// Mitsubishi GX Works2 project: 미니프로젝트 합본   PLC: Q03UDV

PROGRAM MAIN
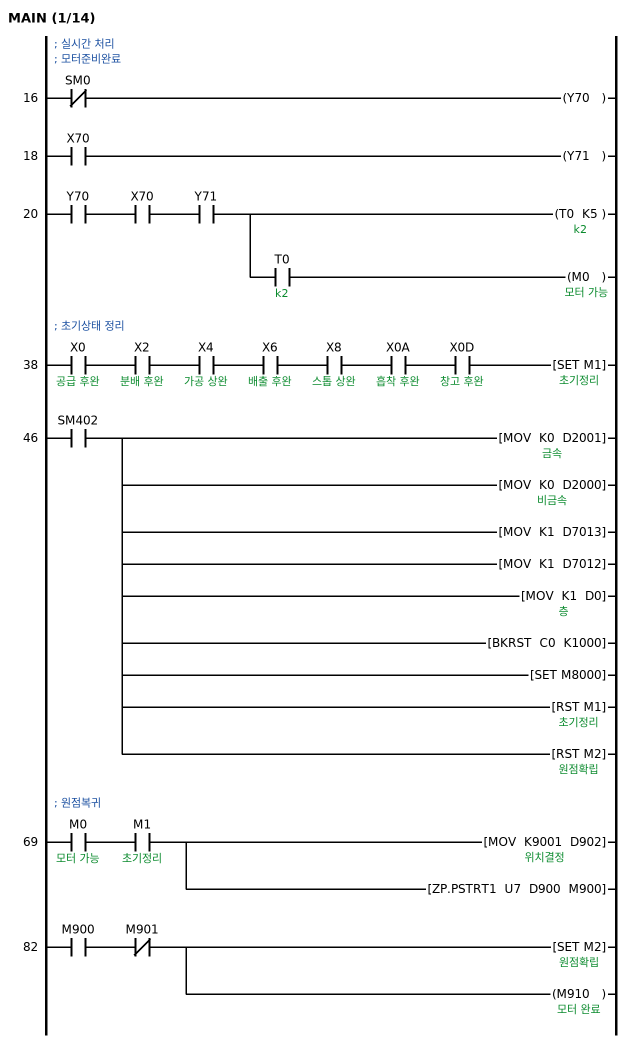
; 실시간 처리
; 모터준비완료
16    LDI     SM0
      OUT     Y70
18    LD      X70
      OUT     Y71
20    LD      Y70
      AND     X70
      AND     Y71
      OUT     T0 K5  ; k2
      AND     T0  ; k2
      OUT     M0  ; 모터 가능
; 초기상태 정리
38    LD      X0  ; 공급 후완
      AND     X2  ; 분배 후완
      AND     X4  ; 가공 상완
      AND     X6  ; 배출 후완
      AND     X8  ; 스톱 상완
      AND     X0A  ; 흡착 후완
      AND     X0D  ; 창고 후완
      SET     M1  ; 초기정리
46    LD      SM402
      MOV     K0 D2001  ; 금속
      MOV     K0 D2000  ; 비금속
      MOV     K1 D7013
      MOV     K1 D7012
      MOV     K1 D0  ; 층
      BKRST   C0 K1000
      SET     M8000
      RST     M1  ; 초기정리
      RST     M2  ; 원점확립
; 원점복귀
69    LD      M0  ; 모터 가능
      AND     M1  ; 초기정리
      MOV     K9001 D902  ; 위치결정
      ZP.PSTRT1 U7 D900 M900
82    LD      M900
      ANI     M901
      SET     M2  ; 원점확립
      OUT     M910  ; 모터 완료
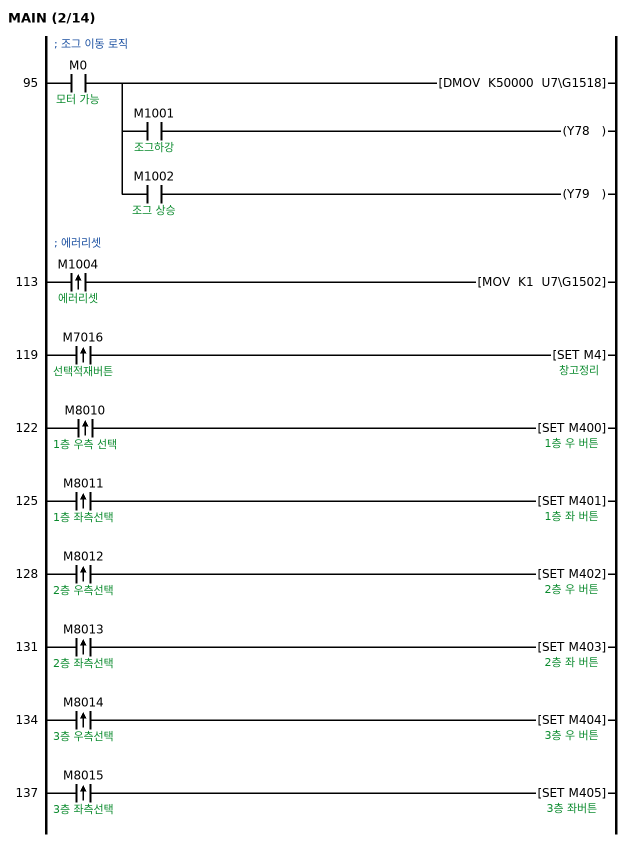
; 조그 이동 로직
95    LD      M0  ; 모터 가능
      DMOV    K50000 U7\G1518
      MPS
      AND     M1001  ; 조그하강
      OUT     Y78
      MPP
      AND     M1002  ; 조그 상승
      OUT     Y79
; 에러리셋
113   LDP     M1004  ; 에러리셋
      MOV     K1 U7\G1502
119   LDP     M7016  ; 선택적재버튼
      SET     M4  ; 창고정리
122   LDP     M8010  ; 1층 우측 선택
      SET     M400  ; 1층 우 버튼
125   LDP     M8011  ; 1층 좌측선택
      SET     M401  ; 1층 좌 버튼
128   LDP     M8012  ; 2층 우측선택
      SET     M402  ; 2층 우 버튼
131   LDP     M8013  ; 2층 좌측선택
      SET     M403  ; 2층 좌 버튼
134   LDP     M8014  ; 3층 우측선택
      SET     M404  ; 3층 우 버튼
137   LDP     M8015  ; 3층 좌측선택
      SET     M405  ; 3층 좌버튼
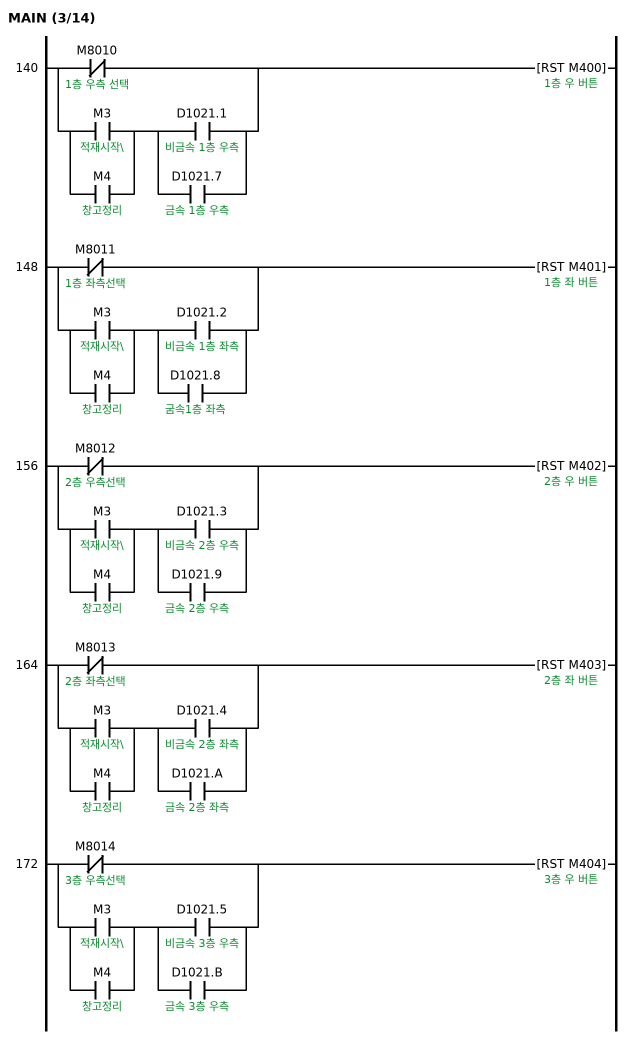
140   LDI     M8010  ; 1층 우측 선택
      LD      M3  ; 적재시작\
      OR      M4  ; 창고정리
      LD      D1021.1  ; 비금속 1층 우측
      OR      D1021.7  ; 금속 1층 우측
      ANB
      ORB
      RST     M400  ; 1층 우 버튼
148   LDI     M8011  ; 1층 좌측선택
      LD      M3  ; 적재시작\
      OR      M4  ; 창고정리
      LD      D1021.2  ; 비금속 1층 좌측
      OR      D1021.8  ; 굼속1층 좌측
      ANB
      ORB
      RST     M401  ; 1층 좌 버튼
156   LDI     M8012  ; 2층 우측선택
      LD      M3  ; 적재시작\
      OR      M4  ; 창고정리
      LD      D1021.3  ; 비금속 2층 우측
      OR      D1021.9  ; 금속 2층 우측
      ANB
      ORB
      RST     M402  ; 2층 우 버튼
164   LDI     M8013  ; 2층 좌측선택
      LD      M3  ; 적재시작\
      OR      M4  ; 창고정리
      LD      D1021.4  ; 비금속 2층 좌측
      OR      D1021.A  ; 금속 2층 좌측
      ANB
      ORB
      RST     M403  ; 2층 좌 버튼
172   LDI     M8014  ; 3층 우측선택
      LD      M3  ; 적재시작\
      OR      M4  ; 창고정리
      LD      D1021.5  ; 비금속 3층 우측
      OR      D1021.B  ; 금속 3층 우측
      ANB
      ORB
      RST     M404  ; 3층 우 버튼
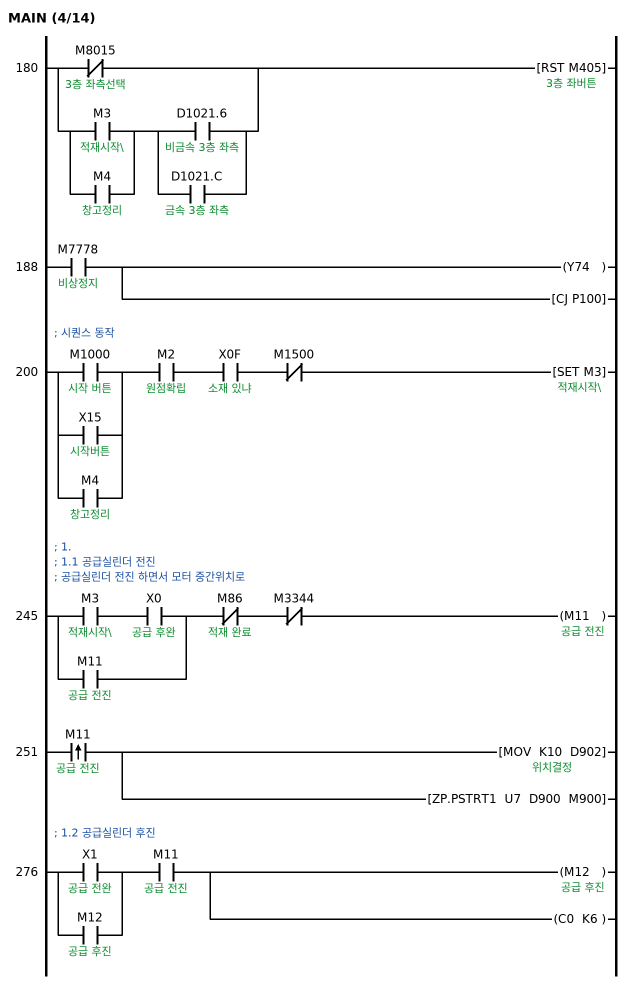
180   LDI     M8015  ; 3층 좌측선택
      LD      M3  ; 적재시작\
      OR      M4  ; 창고정리
      LD      D1021.6  ; 비금속 3층 좌측
      OR      D1021.C  ; 금속 3층 좌측
      ANB
      ORB
      RST     M405  ; 3층 좌버튼
188   LD      M7778  ; 비상정지
      OUT     Y74
      CJ      P100
; 시퀀스 동작
200   LD      M1000  ; 시작 버튼
      OR      X15  ; 시작버튼
      OR      M4  ; 창고정리
      AND     M2  ; 원점확립
      AND     X0F  ; 소재 있냐
      ANI     M1500
      SET     M3  ; 적재시작\
; 1.
; 1.1 공급실린더 전진
; 공급실린더 전진 하면서 모터 중간위치로
245   LD      M3  ; 적재시작\
      AND     X0  ; 공급 후완
      OR      M11  ; 공급 전진
      ANI     M86  ; 적재 완료
      ANI     M3344
      OUT     M11  ; 공급 전진
251   LDP     M11  ; 공급 전진
      MOV     K10 D902
      ZP.PSTRT1 U7 D900 M900
; 1.2 공급실린더 후진
276   LD      X1  ; 공급 전완
      OR      M12  ; 공급 후진
      AND     M11  ; 공급 전진
      OUT     M12  ; 공급 후진
      OUT     C0 K6
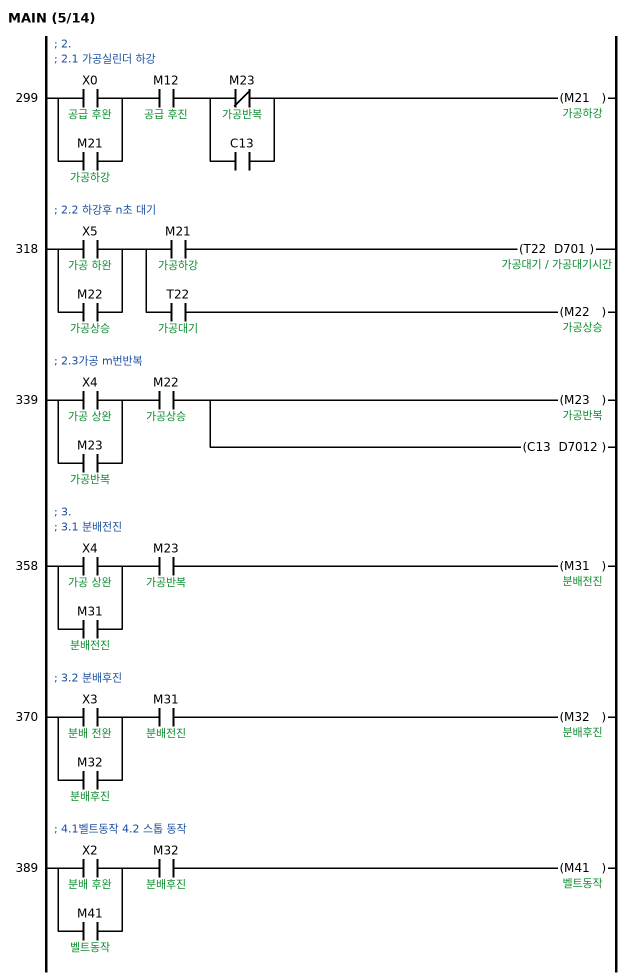
; 2.
; 2.1 가공실린더 하강
299   LD      X0  ; 공급 후완
      OR      M21  ; 가공하강
      AND     M12  ; 공급 후진
      LDI     M23  ; 가공반복
      OR      C13
      ANB
      OUT     M21  ; 가공하강
; 2.2 하강후 n초 대기
318   LD      X5  ; 가공 하완
      OR      M22  ; 가공상승
      MPS
      AND     M21  ; 가공하강
      OUT     T22 D701  ; 가공대기 / 가공대기시간
      MPP
      AND     T22  ; 가공대기
      OUT     M22  ; 가공상승
; 2.3가공 m번반복
339   LD      X4  ; 가공 상완
      OR      M23  ; 가공반복
      AND     M22  ; 가공상승
      OUT     M23  ; 가공반복
      OUT     C13 D7012
; 3.
; 3.1 분배전진
358   LD      X4  ; 가공 상완
      OR      M31  ; 분배전진
      AND     M23  ; 가공반복
      OUT     M31  ; 분배전진
; 3.2 분배후진
370   LD      X3  ; 분배 전완
      OR      M32  ; 분배후진
      AND     M31  ; 분배전진
      OUT     M32  ; 분배후진
; 4.1벨트동작 4.2 스톱 동작
389   LD      X2  ; 분배 후완
      OR      M41  ; 벨트동작
      AND     M32  ; 분배후진
      OUT     M41  ; 벨트동작
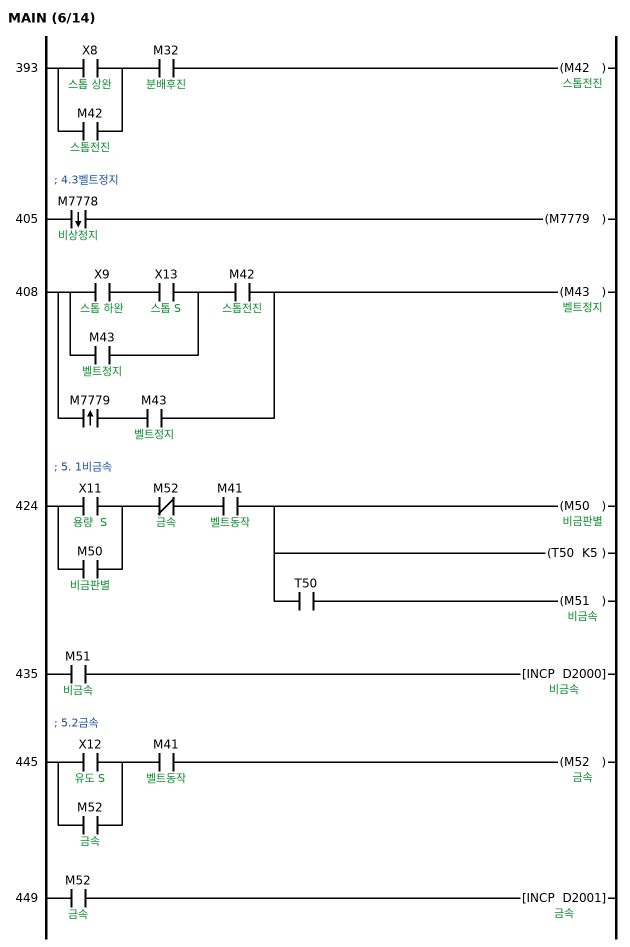
393   LD      X8  ; 스톱 상완
      OR      M42  ; 스톱전진
      AND     M32  ; 분배후진
      OUT     M42  ; 스톱전진
; 4.3벨트정지
405   LDF     M7778  ; 비상정지
      OUT     M7779
408   LD      X9  ; 스톱 하완
      AND     X13  ; 스톱 S
      OR      M43  ; 벨트정지
      AND     M42  ; 스톱전진
      LDP     M7779
      AND     M43  ; 벨트정지
      ORB
      OUT     M43  ; 벨트정지
; 5. 1비금속
424   LD      X11  ; 용량  S
      OR      M50  ; 비금판별
      ANI     M52  ; 금속
      AND     M41  ; 벨트동작
      OUT     M50  ; 비금판별
      OUT     T50 K5
      AND     T50
      OUT     M51  ; 비금속
435   LD      M51  ; 비금속
      INCP    D2000
; 5.2금속
445   LD      X12  ; 유도 S
      OR      M52  ; 금속
      AND     M41  ; 벨트동작
      OUT     M52  ; 금속
449   LD      M52  ; 금속
      INCP    D2001
      P100
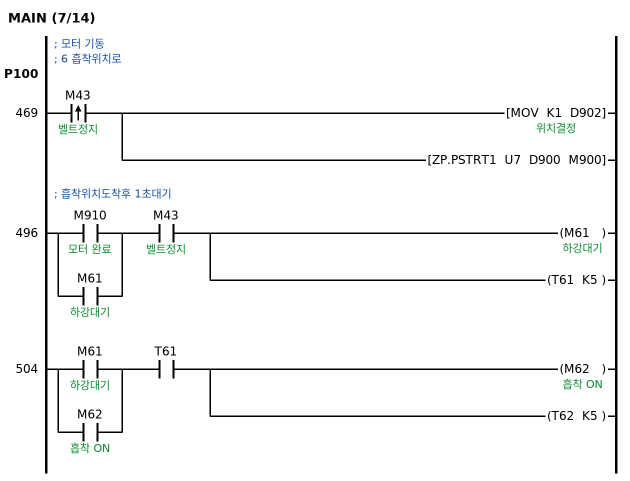
; 모터 기동
; 6 흡착위치로
469   LDP     M43  ; 벨트정지
      MOV     K1 D902
      ZP.PSTRT1 U7 D900 M900
; 흡착위치도착후 1초대기
496   LD      M910  ; 모터 완료
      OR      M61  ; 하강대기
      AND     M43  ; 벨트정지
      OUT     M61  ; 하강대기
      OUT     T61 K5
504   LD      M61  ; 하강대기
      OR      M62  ; 흡착 ON
      AND     T61
      OUT     M62  ; 흡착 ON
      OUT     T62 K5
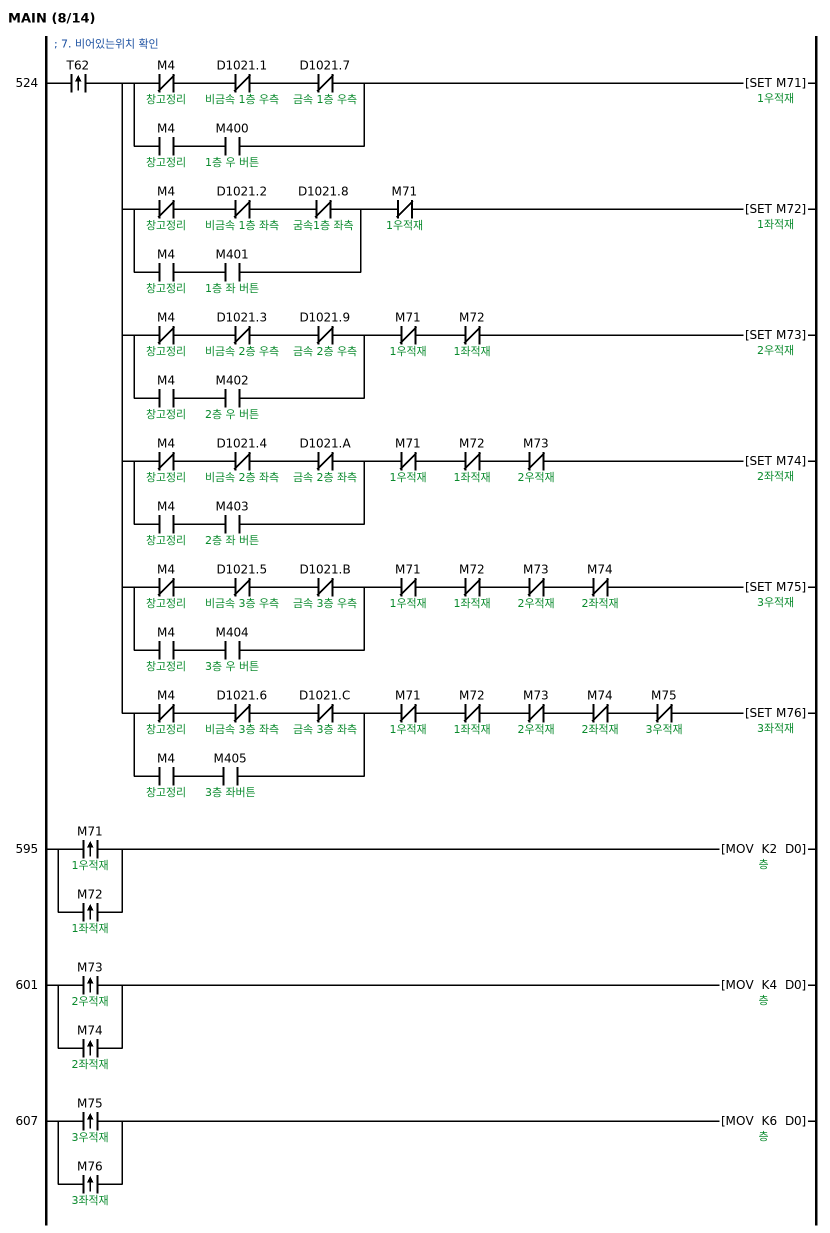
; 7. 비어있는위치 확인
524   LDP     T62
      MPS
      LDI     M4  ; 창고정리
      ANI     D1021.1  ; 비금속 1층 우측
      ANI     D1021.7  ; 금속 1층 우측
      LD      M4  ; 창고정리
      AND     M400  ; 1층 우 버튼
      ORB
      ANB
      SET     M71  ; 1우적재
      MRD
      LDI     M4  ; 창고정리
      ANI     D1021.2  ; 비금속 1층 좌측
      ANI     D1021.8  ; 굼속1층 좌측
      LD      M4  ; 창고정리
      AND     M401  ; 1층 좌 버튼
      ORB
      ANB
      ANI     M71  ; 1우적재
      SET     M72  ; 1좌적재
      MRD
      LDI     M4  ; 창고정리
      ANI     D1021.3  ; 비금속 2층 우측
      ANI     D1021.9  ; 금속 2층 우측
      LD      M4  ; 창고정리
      AND     M402  ; 2층 우 버튼
      ORB
      ANB
      ANI     M71  ; 1우적재
      ANI     M72  ; 1좌적재
      SET     M73  ; 2우적재
      MRD
      LDI     M4  ; 창고정리
      ANI     D1021.4  ; 비금속 2층 좌측
      ANI     D1021.A  ; 금속 2층 좌측
      LD      M4  ; 창고정리
      AND     M403  ; 2층 좌 버튼
      ORB
      ANB
      ANI     M71  ; 1우적재
      ANI     M72  ; 1좌적재
      ANI     M73  ; 2우적재
      SET     M74  ; 2좌적재
      MRD
      LDI     M4  ; 창고정리
      ANI     D1021.5  ; 비금속 3층 우측
      ANI     D1021.B  ; 금속 3층 우측
      LD      M4  ; 창고정리
      AND     M404  ; 3층 우 버튼
      ORB
      ANB
      ANI     M71  ; 1우적재
      ANI     M72  ; 1좌적재
      ANI     M73  ; 2우적재
      ANI     M74  ; 2좌적재
      SET     M75  ; 3우적재
      MPP
      LDI     M4  ; 창고정리
      ANI     D1021.6  ; 비금속 3층 좌측
      ANI     D1021.C  ; 금속 3층 좌측
      LD      M4  ; 창고정리
      AND     M405  ; 3층 좌버튼
      ORB
      ANB
      ANI     M71  ; 1우적재
      ANI     M72  ; 1좌적재
      ANI     M73  ; 2우적재
      ANI     M74  ; 2좌적재
      ANI     M75  ; 3우적재
      SET     M76  ; 3좌적재
595   LDP     M71  ; 1우적재
      ORP     M72  ; 1좌적재
      MOV     K2 D0
601   LDP     M73  ; 2우적재
      ORP     M74  ; 2좌적재
      MOV     K4 D0
607   LDP     M75  ; 3우적재
      ORP     M76  ; 3좌적재
      MOV     K6 D0
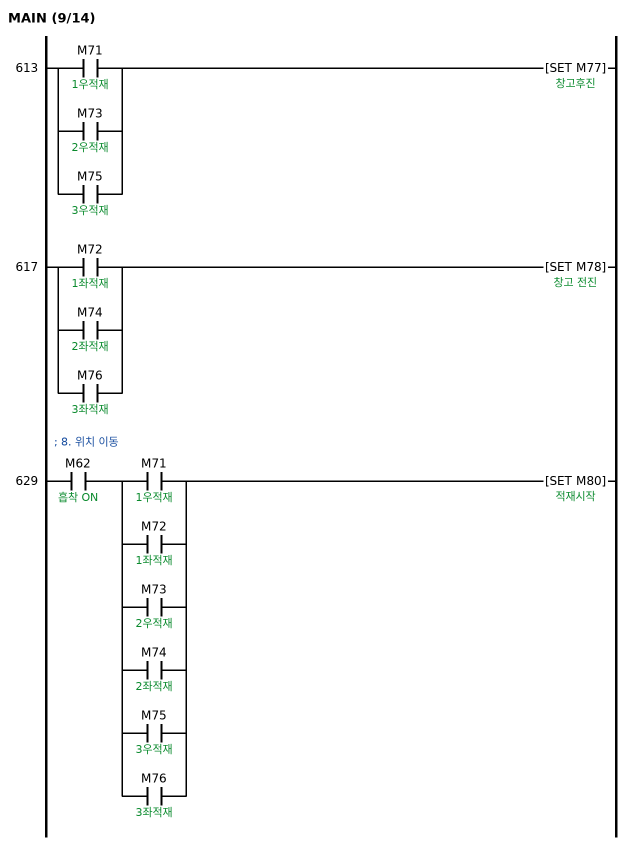
613   LD      M71  ; 1우적재
      OR      M73  ; 2우적재
      OR      M75  ; 3우적재
      SET     M77  ; 창고후진
617   LD      M72  ; 1좌적재
      OR      M74  ; 2좌적재
      OR      M76  ; 3좌적재
      SET     M78  ; 창고 전진
; 8. 위치 이동
629   LD      M62  ; 흡착 ON
      LD      M71  ; 1우적재
      OR      M72  ; 1좌적재
      OR      M73  ; 2우적재
      OR      M74  ; 2좌적재
      OR      M75  ; 3우적재
      OR      M76  ; 3좌적재
      ANB
      SET     M80  ; 적재시작
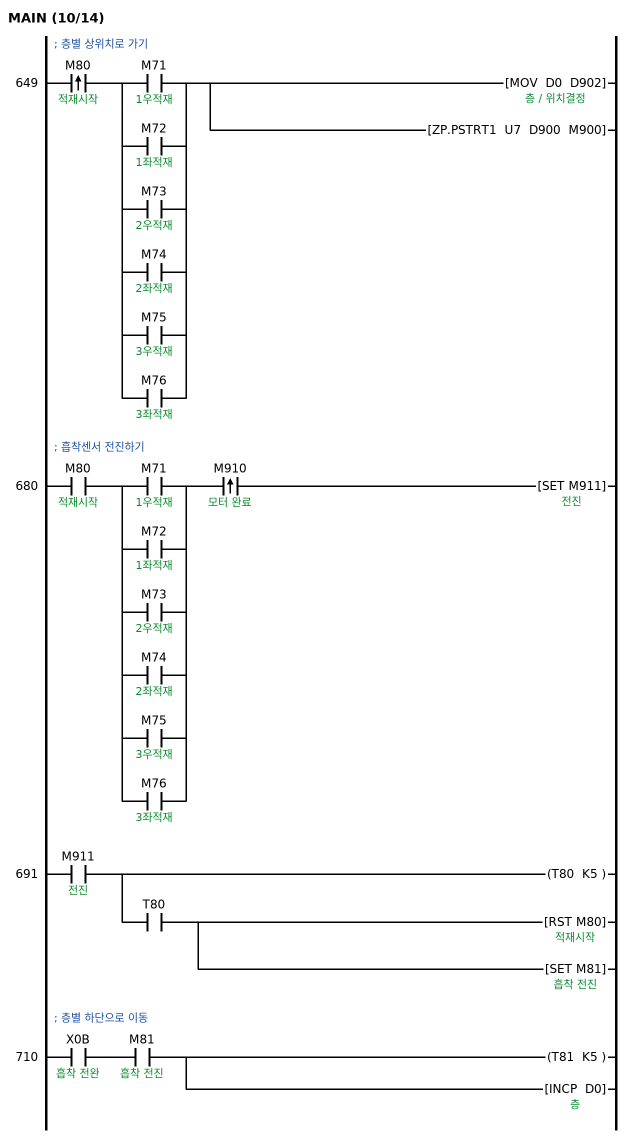
; 층별 상위치로 가기
649   LDP     M80  ; 적재시작
      LD      M71  ; 1우적재
      OR      M72  ; 1좌적재
      OR      M73  ; 2우적재
      OR      M74  ; 2좌적재
      OR      M75  ; 3우적재
      OR      M76  ; 3좌적재
      ANB
      MOV     D0 D902
      ZP.PSTRT1 U7 D900 M900
; 흡착센서 전진하기
680   LD      M80  ; 적재시작
      LD      M71  ; 1우적재
      OR      M72  ; 1좌적재
      OR      M73  ; 2우적재
      OR      M74  ; 2좌적재
      OR      M75  ; 3우적재
      OR      M76  ; 3좌적재
      ANB
      ANDP    M910  ; 모터 완료
      SET     M911  ; 전진
691   LD      M911  ; 전진
      OUT     T80 K5
      AND     T80
      RST     M80  ; 적재시작
      SET     M81  ; 흡착 전진
; 층별 하단으로 이동
710   LD      X0B  ; 흡착 전완
      AND     M81  ; 흡착 전진
      OUT     T81 K5
      INCP    D0
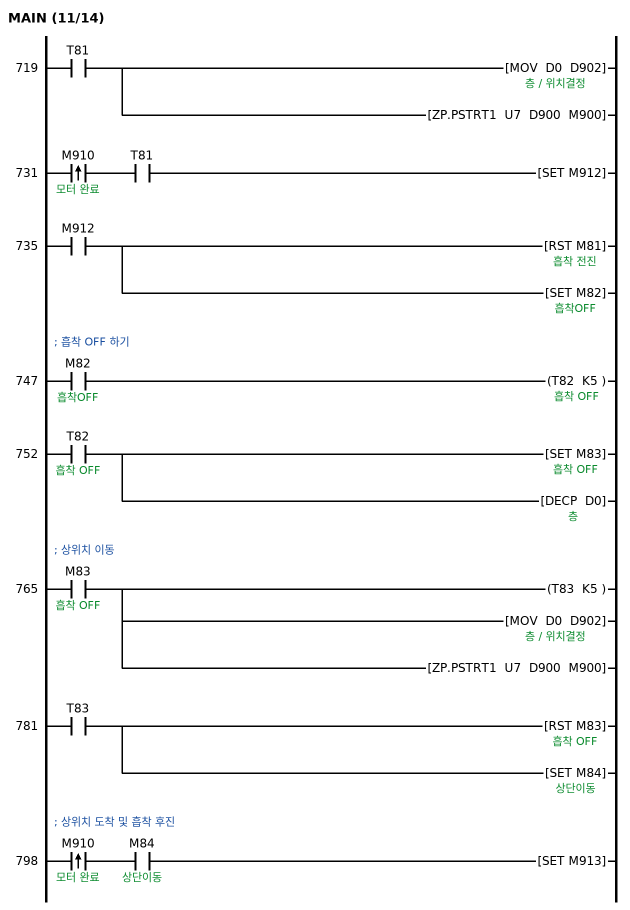
719   LD      T81
      MOV     D0 D902
      ZP.PSTRT1 U7 D900 M900
731   LDP     M910  ; 모터 완료
      AND     T81
      SET     M912
735   LD      M912
      RST     M81  ; 흡착 전진
      SET     M82  ; 흡착OFF
; 흡착 OFF 하기
747   LD      M82  ; 흡착OFF
      OUT     T82 K5  ; 흡착 OFF
752   LD      T82  ; 흡착 OFF
      SET     M83  ; 흡착 OFF
      DECP    D0
; 상위치 이동
765   LD      M83  ; 흡착 OFF
      OUT     T83 K5
      MOV     D0 D902
      ZP.PSTRT1 U7 D900 M900
781   LD      T83
      RST     M83  ; 흡착 OFF
      SET     M84  ; 상단이동
; 상위치 도착 및 흡착 후진
798   LDP     M910  ; 모터 완료
      AND     M84  ; 상단이동
      SET     M913
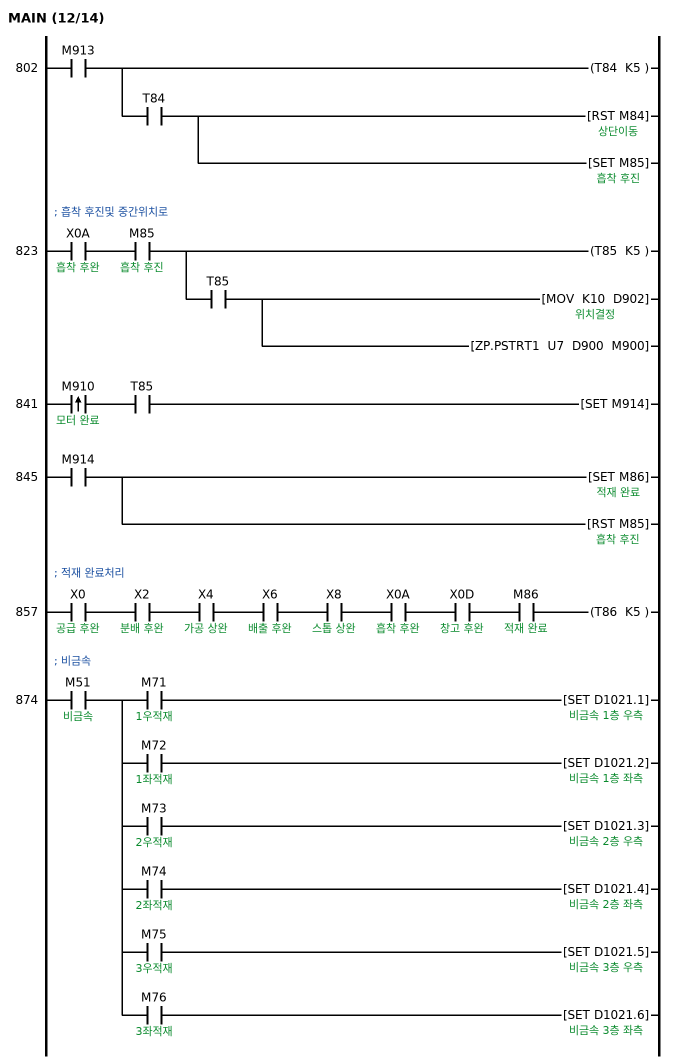
802   LD      M913
      OUT     T84 K5
      AND     T84
      RST     M84  ; 상단이동
      SET     M85  ; 흡착 후진
; 흡착 후진및 중간위치로
823   LD      X0A  ; 흡착 후완
      AND     M85  ; 흡착 후진
      OUT     T85 K5
      AND     T85
      MOV     K10 D902
      ZP.PSTRT1 U7 D900 M900
841   LDP     M910  ; 모터 완료
      AND     T85
      SET     M914
845   LD      M914
      SET     M86  ; 적재 완료
      RST     M85  ; 흡착 후진
; 적재 완료처리
857   LD      X0  ; 공급 후완
      AND     X2  ; 분배 후완
      AND     X4  ; 가공 상완
      AND     X6  ; 배출 후완
      AND     X8  ; 스톱 상완
      AND     X0A  ; 흡착 후완
      AND     X0D  ; 창고 후완
      AND     M86  ; 적재 완료
      OUT     T86 K5
; 비금속
874   LD      M51  ; 비금속
      MPS
      AND     M71  ; 1우적재
      SET     D1021.1  ; 비금속 1층 우측
      MRD
      AND     M72  ; 1좌적재
      SET     D1021.2  ; 비금속 1층 좌측
      MRD
      AND     M73  ; 2우적재
      SET     D1021.3  ; 비금속 2층 우측
      MRD
      AND     M74  ; 2좌적재
      SET     D1021.4  ; 비금속 2층 좌측
      MRD
      AND     M75  ; 3우적재
      SET     D1021.5  ; 비금속 3층 우측
      MPP
      AND     M76  ; 3좌적재
      SET     D1021.6  ; 비금속 3층 좌측
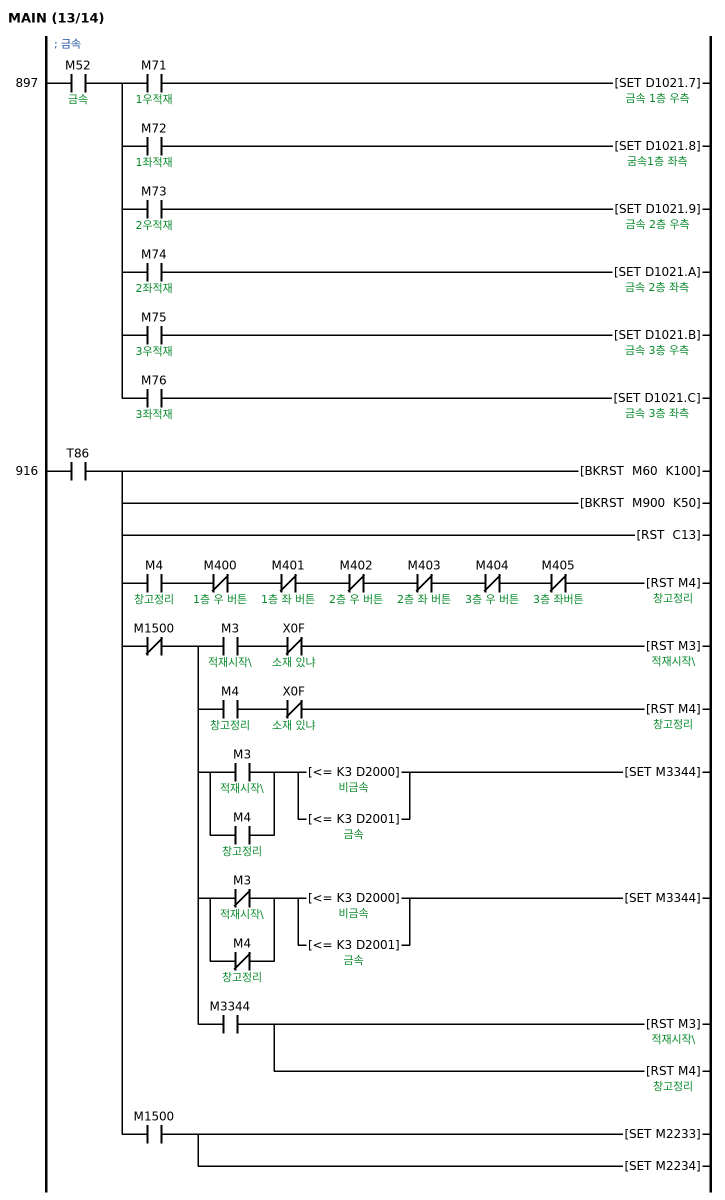
; 금속
897   LD      M52  ; 금속
      MPS
      AND     M71  ; 1우적재
      SET     D1021.7  ; 금속 1층 우측
      MRD
      AND     M72  ; 1좌적재
      SET     D1021.8  ; 굼속1층 좌측
      MRD
      AND     M73  ; 2우적재
      SET     D1021.9  ; 금속 2층 우측
      MRD
      AND     M74  ; 2좌적재
      SET     D1021.A  ; 금속 2층 좌측
      MRD
      AND     M75  ; 3우적재
      SET     D1021.B  ; 금속 3층 우측
      MPP
      AND     M76  ; 3좌적재
      SET     D1021.C  ; 금속 3층 좌측
916   LD      T86
      BKRST   M60 K100
      BKRST   M900 K50
      RST     C13
      MPS
      AND     M4  ; 창고정리
      ANI     M400  ; 1층 우 버튼
      ANI     M401  ; 1층 좌 버튼
      ANI     M402  ; 2층 우 버튼
      ANI     M403  ; 2층 좌 버튼
      ANI     M404  ; 3층 우 버튼
      ANI     M405  ; 3층 좌버튼
      RST     M4  ; 창고정리
      MRD
      ANI     M1500
      MPS
      AND     M3  ; 적재시작\
      ANI     X0F  ; 소재 있냐
      RST     M3  ; 적재시작\
      MRD
      AND     M4  ; 창고정리
      ANI     X0F  ; 소재 있냐
      RST     M4  ; 창고정리
      MRD
      LD      M3  ; 적재시작\
      OR      M4  ; 창고정리
      ANB
      LD<=    K3 D2000  ; 비금속
      OR<=    K3 D2001  ; 금속
      ANB
      SET     M3344
      MRD
      LDI     M3  ; 적재시작\
      ORI     M4  ; 창고정리
      ANB
      LD<=    K3 D2000  ; 비금속
      OR<=    K3 D2001  ; 금속
      ANB
      SET     M3344
      MPP
      AND     M3344
      RST     M3  ; 적재시작\
      RST     M4  ; 창고정리
      MPP
      AND     M1500
      SET     M2233
      SET     M2234
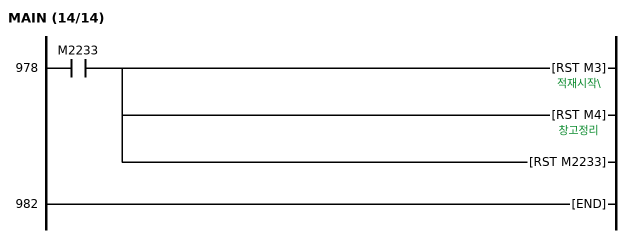
978   LD      M2233
      RST     M3  ; 적재시작\
      RST     M4  ; 창고정리
      RST     M2233
982   END
END_PROGRAM

PROGRAM OUTPUT
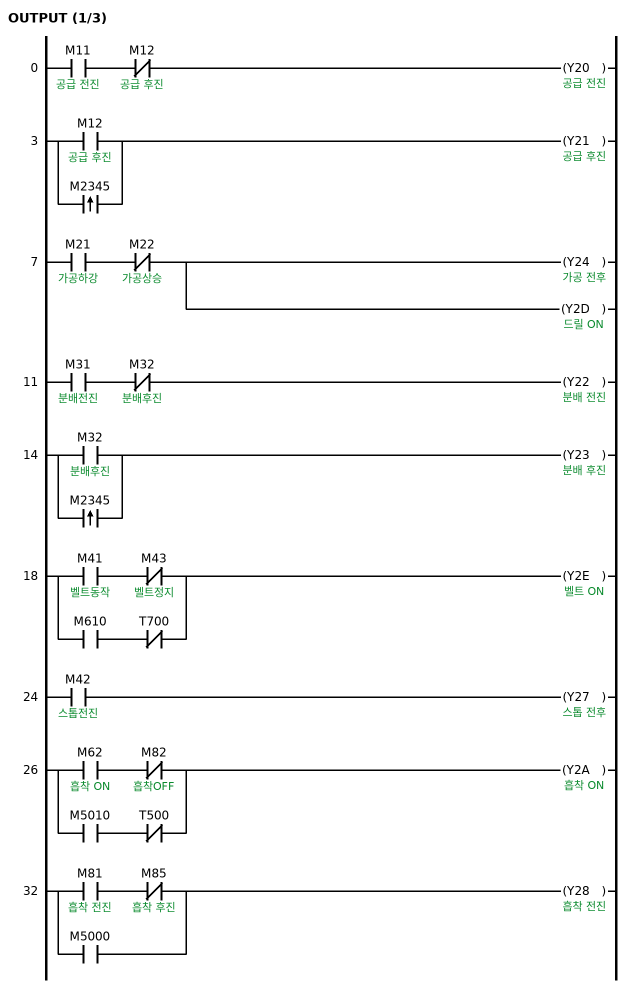
0     LD      M11  ; 공급 전진
      ANI     M12  ; 공급 후진
      OUT     Y20  ; 공급 전진
3     LD      M12  ; 공급 후진
      ORP     M2345
      OUT     Y21  ; 공급 후진
7     LD      M21  ; 가공하강
      ANI     M22  ; 가공상승
      OUT     Y24  ; 가공 전후
      OUT     Y2D  ; 드릴 ON
11    LD      M31  ; 분배전진
      ANI     M32  ; 분배후진
      OUT     Y22  ; 분배 전진
14    LD      M32  ; 분배후진
      ORP     M2345
      OUT     Y23  ; 분배 후진
18    LD      M41  ; 벨트동작
      ANI     M43  ; 벨트정지
      LD      M610
      ANI     T700
      ORB
      OUT     Y2E  ; 벨트 ON
24    LD      M42  ; 스톱전진
      OUT     Y27  ; 스톱 전후
26    LD      M62  ; 흡착 ON
      ANI     M82  ; 흡착OFF
      LD      M5010
      ANI     T500
      ORB
      OUT     Y2A  ; 흡착 ON
32    LD      M81  ; 흡착 전진
      ANI     M85  ; 흡착 후진
      OR      M5000
      OUT     Y28  ; 흡착 전진
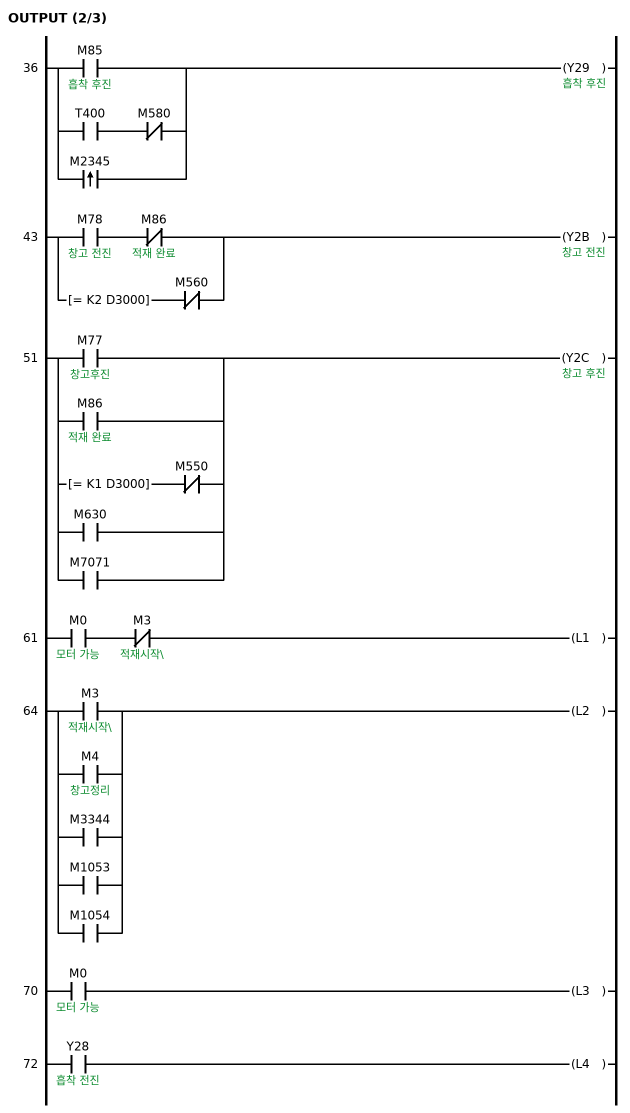
36    LD      M85  ; 흡착 후진
      LD      T400
      ANI     M580
      ORB
      ORP     M2345
      OUT     Y29  ; 흡착 후진
43    LD      M78  ; 창고 전진
      ANI     M86  ; 적재 완료
      LD=     K2 D3000
      ANI     M560
      ORB
      OUT     Y2B  ; 창고 전진
51    LD      M77  ; 창고후진
      OR      M86  ; 적재 완료
      LD=     K1 D3000
      ANI     M550
      ORB
      OR      M630
      OR      M7071
      OUT     Y2C  ; 창고 후진
61    LD      M0  ; 모터 가능
      ANI     M3  ; 적재시작\
      OUT     L1
64    LD      M3  ; 적재시작\
      OR      M4  ; 창고정리
      OR      M3344
      OR      M1053
      OR      M1054
      OUT     L2
70    LD      M0  ; 모터 가능
      OUT     L3
72    LD      Y28  ; 흡착 전진
      OUT     L4
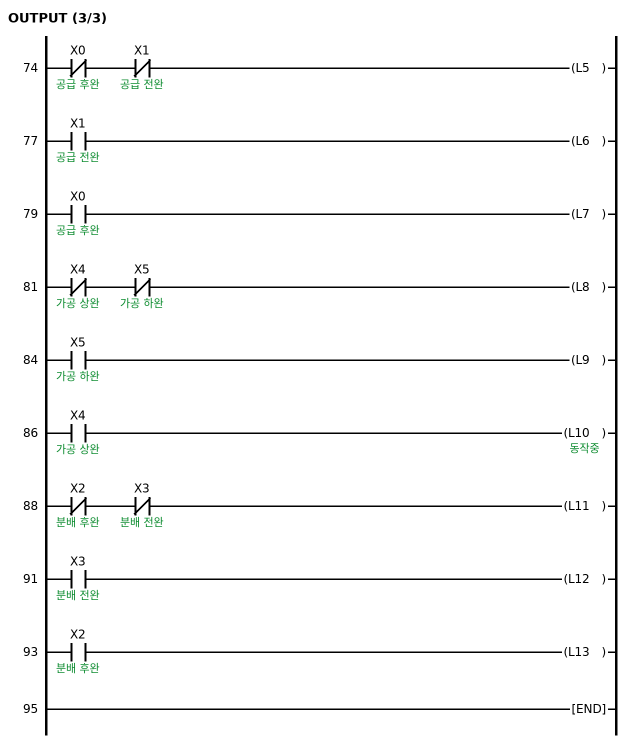
74    LDI     X0  ; 공급 후완
      ANI     X1  ; 공급 전완
      OUT     L5
77    LD      X1  ; 공급 전완
      OUT     L6
79    LD      X0  ; 공급 후완
      OUT     L7
81    LDI     X4  ; 가공 상완
      ANI     X5  ; 가공 하완
      OUT     L8
84    LD      X5  ; 가공 하완
      OUT     L9
86    LD      X4  ; 가공 상완
      OUT     L10  ; 동작중
88    LDI     X2  ; 분배 후완
      ANI     X3  ; 분배 전완
      OUT     L11
91    LD      X3  ; 분배 전완
      OUT     L12
93    LD      X2  ; 분배 후완
      OUT     L13
95    END
END_PROGRAM

PROGRAM HMI
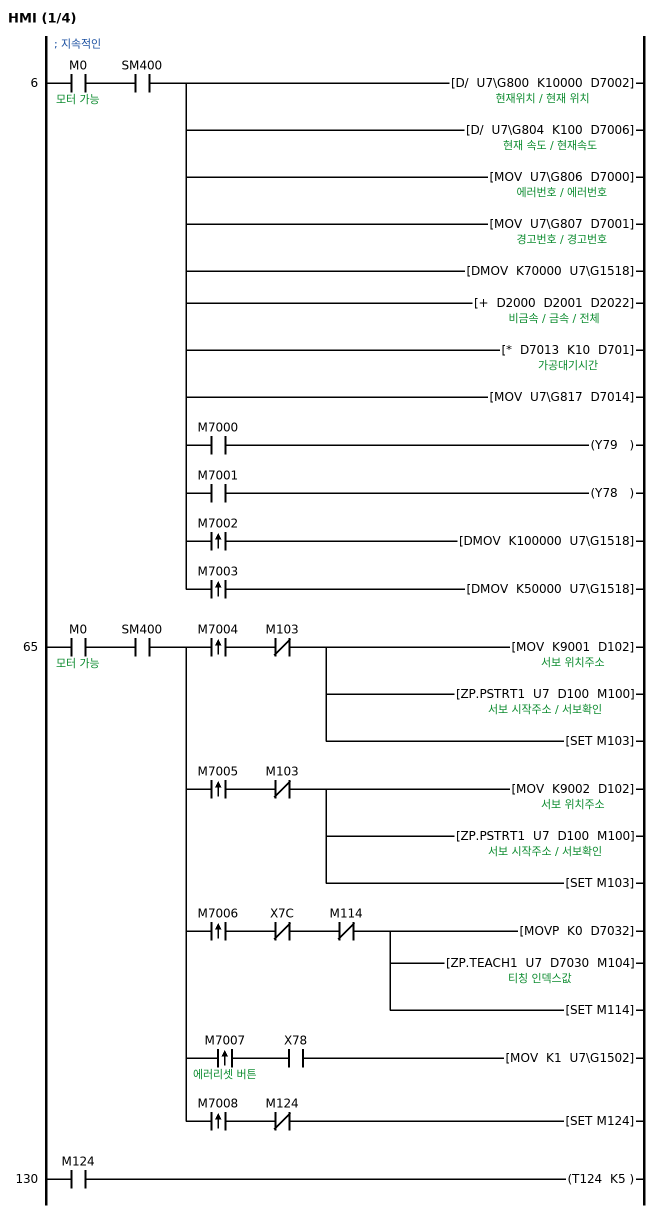
; 지속적인
6     LD      M0  ; 모터 가능
      AND     SM400
      D/      U7\G800 K10000 D7002  ; 현재위치 / 현재 위치
      D/      U7\G804 K100 D7006  ; 현재 속도 / 현재속도
      MOV     U7\G806 D7000  ; 에러번호 / 에러번호
      MOV     U7\G807 D7001  ; 경고번호 / 경고번호
      DMOV    K70000 U7\G1518
      +       D2000 D2001 D2022  ; 비금속 / 금속 / 전체
      *       D7013 K10 D701  ; 가공대기시간
      MOV     U7\G817 D7014
      MPS
      AND     M7000
      OUT     Y79
      MRD
      AND     M7001
      OUT     Y78
      MRD
      ANDP    M7002
      DMOV    K100000 U7\G1518
      MPP
      ANDP    M7003
      DMOV    K50000 U7\G1518
65    LD      M0  ; 모터 가능
      AND     SM400
      MPS
      ANDP    M7004
      ANI     M103
      MOV     K9001 D102  ; 서보 위치주소
      ZP.PSTRT1 U7 D100 M100  ; 서보 시작주소 / 서보확인
      SET     M103
      MRD
      ANDP    M7005
      ANI     M103
      MOV     K9002 D102
      ZP.PSTRT1 U7 D100 M100
      SET     M103
      MRD
      ANDP    M7006
      ANI     X7C
      ANI     M114
      MOVP    K0 D7032
      ZP.TEACH1 U7 D7030 M104  ; 티칭 인덱스값
      SET     M114
      MRD
      ANDP    M7007  ; 에러리셋 버튼
      AND     X78
      MOV     K1 U7\G1502
      MPP
      ANDP    M7008
      ANI     M124
      SET     M124
130   LD      M124
      OUT     T124 K5
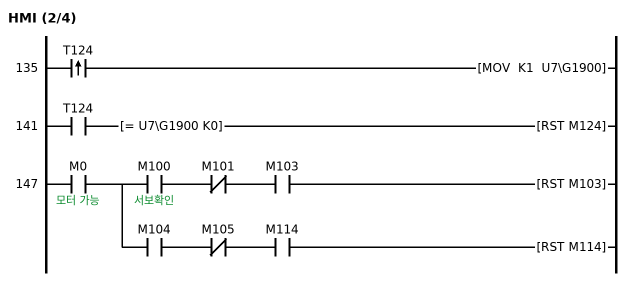
135   LDP     T124
      MOV     K1 U7\G1900
141   LD      T124
      AND=    U7\G1900 K0
      RST     M124
147   LD      M0  ; 모터 가능
      MPS
      AND     M100  ; 서보확인
      ANI     M101
      AND     M103
      RST     M103
      MPP
      AND     M104
      ANI     M105
      AND     M114
      RST     M114
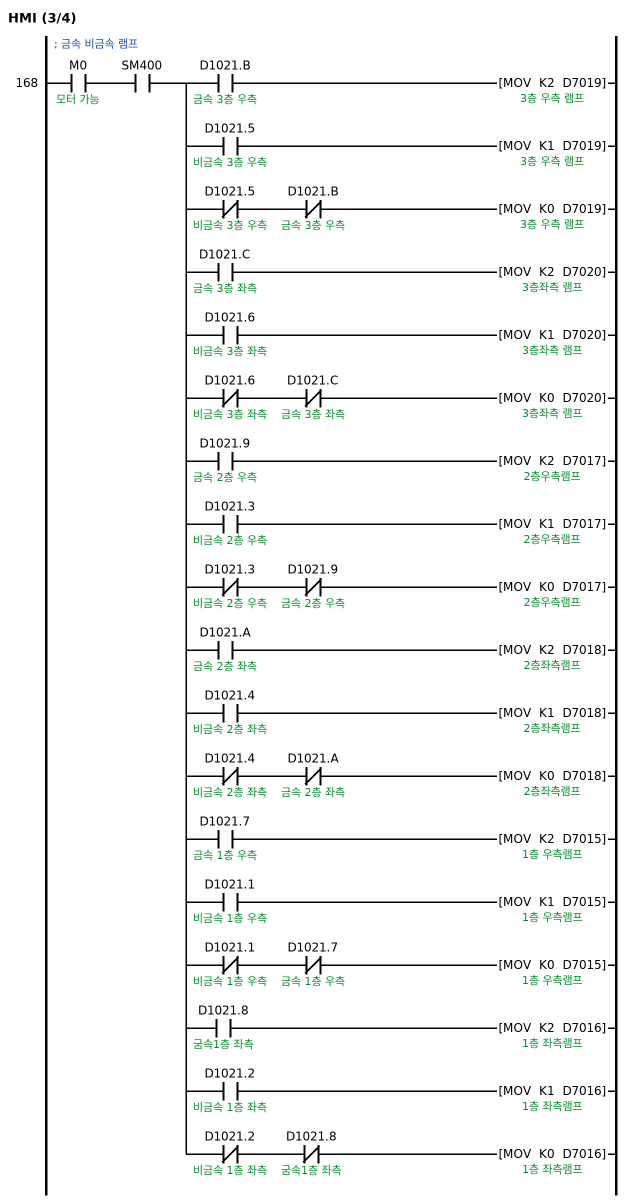
; 금속 비금속 램프
168   LD      M0  ; 모터 가능
      AND     SM400
      MPS
      AND     D1021.B  ; 금속 3층 우측
      MOV     K2 D7019  ; 3층 우측 램프
      MRD
      AND     D1021.5  ; 비금속 3층 우측
      MOV     K1 D7019
      MRD
      ANI     D1021.5  ; 비금속 3층 우측
      ANI     D1021.B  ; 금속 3층 우측
      MOV     K0 D7019
      MRD
      AND     D1021.C  ; 금속 3층 좌측
      MOV     K2 D7020  ; 3층좌측 램프
      MRD
      AND     D1021.6  ; 비금속 3층 좌측
      MOV     K1 D7020
      MRD
      ANI     D1021.6  ; 비금속 3층 좌측
      ANI     D1021.C  ; 금속 3층 좌측
      MOV     K0 D7020
      MRD
      AND     D1021.9  ; 금속 2층 우측
      MOV     K2 D7017  ; 2층우측램프
      MRD
      AND     D1021.3  ; 비금속 2층 우측
      MOV     K1 D7017
      MRD
      ANI     D1021.3  ; 비금속 2층 우측
      ANI     D1021.9  ; 금속 2층 우측
      MOV     K0 D7017
      MRD
      AND     D1021.A  ; 금속 2층 좌측
      MOV     K2 D7018  ; 2층좌측램프
      MRD
      AND     D1021.4  ; 비금속 2층 좌측
      MOV     K1 D7018
      MRD
      ANI     D1021.4  ; 비금속 2층 좌측
      ANI     D1021.A  ; 금속 2층 좌측
      MOV     K0 D7018
      MRD
      AND     D1021.7  ; 금속 1층 우측
      MOV     K2 D7015  ; 1층 우측램프
      MRD
      AND     D1021.1  ; 비금속 1층 우측
      MOV     K1 D7015
      MRD
      ANI     D1021.1  ; 비금속 1층 우측
      ANI     D1021.7  ; 금속 1층 우측
      MOV     K0 D7015
      MRD
      AND     D1021.8  ; 굼속1층 좌측
      MOV     K2 D7016  ; 1층 좌측램프
      MRD
      AND     D1021.2  ; 비금속 1층 좌측
      MOV     K1 D7016
      MPP
      ANI     D1021.2  ; 비금속 1층 좌측
      ANI     D1021.8  ; 굼속1층 좌측
      MOV     K0 D7016
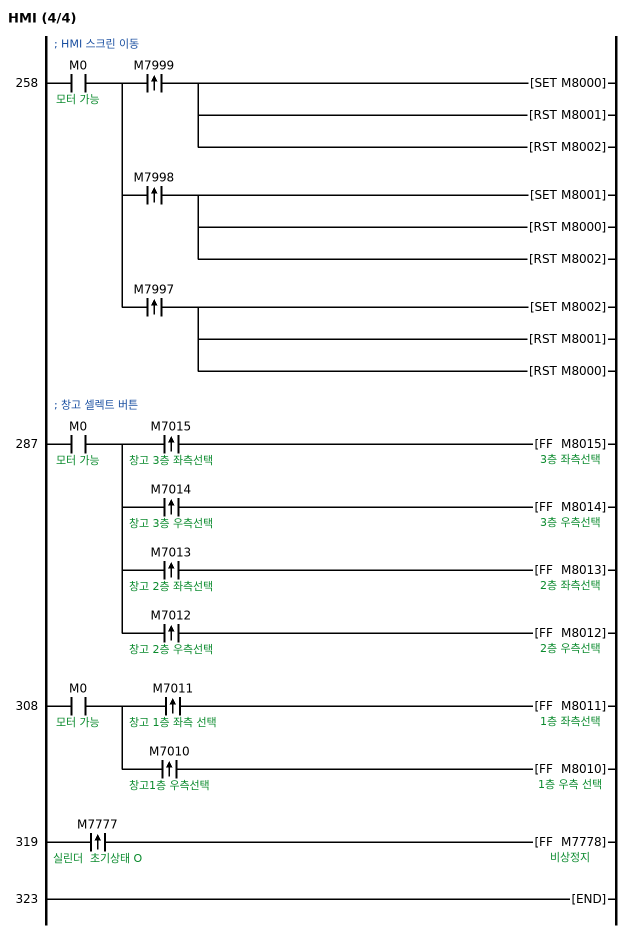
; HMI 스크린 이동
258   LD      M0  ; 모터 가능
      MPS
      ANDP    M7999
      SET     M8000
      RST     M8001
      RST     M8002
      MRD
      ANDP    M7998
      SET     M8001
      RST     M8000
      RST     M8002
      MPP
      ANDP    M7997
      SET     M8002
      RST     M8001
      RST     M8000
; 창고 셀렉트 버튼
287   LD      M0  ; 모터 가능
      MPS
      ANDP    M7015  ; 창고 3층 좌측선택
      FF      M8015  ; 3층 좌측선택
      MRD
      ANDP    M7014  ; 창고 3층 우측선택
      FF      M8014  ; 3층 우측선택
      MRD
      ANDP    M7013  ; 창고 2층 좌측선택
      FF      M8013  ; 2층 좌측선택
      MPP
      ANDP    M7012  ; 창고 2층 우측선택
      FF      M8012  ; 2층 우측선택
308   LD      M0  ; 모터 가능
      MPS
      ANDP    M7011  ; 창고 1층 좌측 선택
      FF      M8011  ; 1층 좌측선택
      MPP
      ANDP    M7010  ; 창고1층 우측선택
      FF      M8010  ; 1층 우측 선택
319   LDP     M7777  ; 실린더  초기상태 O
      FF      M7778  ; 비상정지
323   END
END_PROGRAM

PROGRAM RELEASE
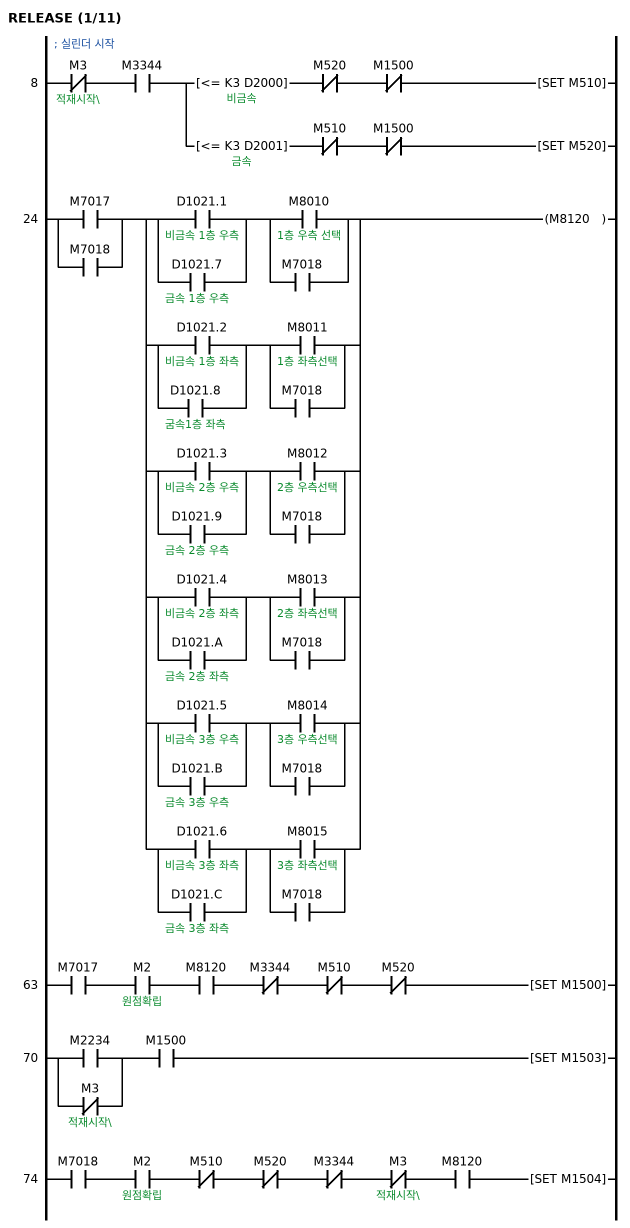
; 실린더 시작
8     LDI     M3  ; 적재시작\
      AND     M3344
      MPS
      AND<=   K3 D2000  ; 비금속
      ANI     M520
      ANI     M1500
      SET     M510
      MPP
      AND<=   K3 D2001  ; 금속
      ANI     M510
      ANI     M1500
      SET     M520
24    LD      M7017
      OR      M7018
      LD      D1021.1  ; 비금속 1층 우측
      OR      D1021.7  ; 금속 1층 우측
      LD      M8010  ; 1층 우측 선택
      OR      M7018
      ANB
      LD      D1021.2  ; 비금속 1층 좌측
      OR      D1021.8  ; 굼속1층 좌측
      LD      M8011  ; 1층 좌측선택
      OR      M7018
      ANB
      ORB
      LD      D1021.3  ; 비금속 2층 우측
      OR      D1021.9  ; 금속 2층 우측
      LD      M8012  ; 2층 우측선택
      OR      M7018
      ANB
      ORB
      LD      D1021.4  ; 비금속 2층 좌측
      OR      D1021.A  ; 금속 2층 좌측
      LD      M8013  ; 2층 좌측선택
      OR      M7018
      ANB
      ORB
      LD      D1021.5  ; 비금속 3층 우측
      OR      D1021.B  ; 금속 3층 우측
      LD      M8014  ; 3층 우측선택
      OR      M7018
      ANB
      ORB
      LD      D1021.6  ; 비금속 3층 좌측
      OR      D1021.C  ; 금속 3층 좌측
      LD      M8015  ; 3층 좌측선택
      OR      M7018
      ANB
      ORB
      ANB
      OUT     M8120
63    LD      M7017
      AND     M2  ; 원점확립
      AND     M8120
      ANI     M3344
      ANI     M510
      ANI     M520
      SET     M1500
70    LD      M2234
      ORI     M3  ; 적재시작\
      AND     M1500
      SET     M1503
74    LD      M7018
      AND     M2  ; 원점확립
      ANI     M510
      ANI     M520
      ANI     M3344
      ANI     M3  ; 적재시작\
      AND     M8120
      SET     M1504
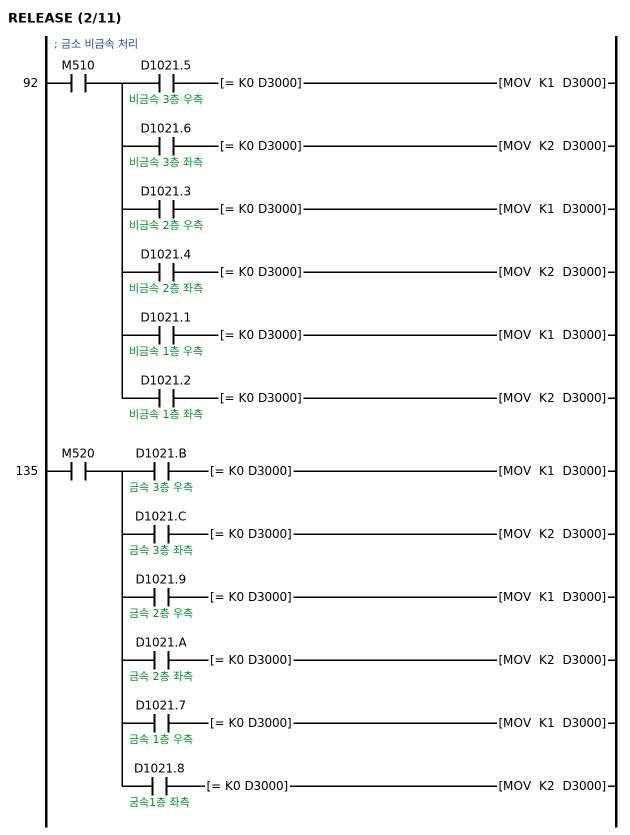
; 금소 비금속 처리
92    LD      M510
      MPS
      AND     D1021.5  ; 비금속 3층 우측
      AND=    K0 D3000
      MOV     K1 D3000
      MRD
      AND     D1021.6  ; 비금속 3층 좌측
      AND=    K0 D3000
      MOV     K2 D3000
      MRD
      AND     D1021.3  ; 비금속 2층 우측
      AND=    K0 D3000
      MOV     K1 D3000
      MRD
      AND     D1021.4  ; 비금속 2층 좌측
      AND=    K0 D3000
      MOV     K2 D3000
      MRD
      AND     D1021.1  ; 비금속 1층 우측
      AND=    K0 D3000
      MOV     K1 D3000
      MPP
      AND     D1021.2  ; 비금속 1층 좌측
      AND=    K0 D3000
      MOV     K2 D3000
135   LD      M520
      MPS
      AND     D1021.B  ; 금속 3층 우측
      AND=    K0 D3000
      MOV     K1 D3000
      MRD
      AND     D1021.C  ; 금속 3층 좌측
      AND=    K0 D3000
      MOV     K2 D3000
      MRD
      AND     D1021.9  ; 금속 2층 우측
      AND=    K0 D3000
      MOV     K1 D3000
      MRD
      AND     D1021.A  ; 금속 2층 좌측
      AND=    K0 D3000
      MOV     K2 D3000
      MRD
      AND     D1021.7  ; 금속 1층 우측
      AND=    K0 D3000
      MOV     K1 D3000
      MPP
      AND     D1021.8  ; 굼속1층 좌측
      AND=    K0 D3000
      MOV     K2 D3000
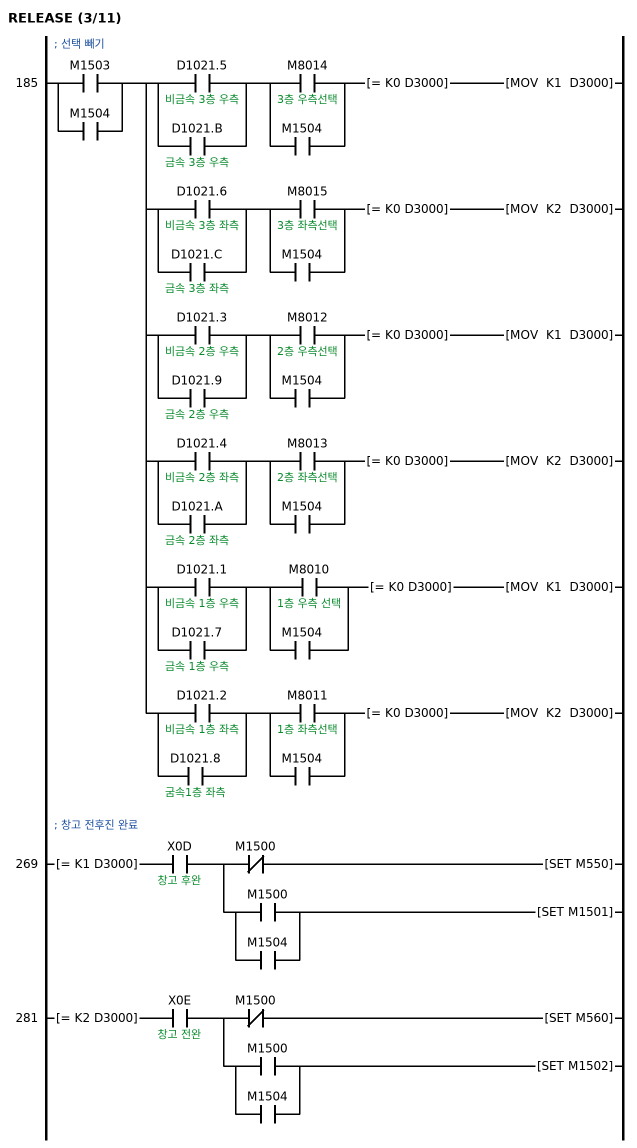
; 선택 빼기
185   LD      M1503
      OR      M1504
      MPS
      LD      D1021.5  ; 비금속 3층 우측
      OR      D1021.B  ; 금속 3층 우측
      ANB
      LD      M8014  ; 3층 우측선택
      OR      M1504
      ANB
      AND=    K0 D3000
      MOV     K1 D3000
      MRD
      LD      D1021.6  ; 비금속 3층 좌측
      OR      D1021.C  ; 금속 3층 좌측
      ANB
      LD      M8015  ; 3층 좌측선택
      OR      M1504
      ANB
      AND=    K0 D3000
      MOV     K2 D3000
      MRD
      LD      D1021.3  ; 비금속 2층 우측
      OR      D1021.9  ; 금속 2층 우측
      ANB
      LD      M8012  ; 2층 우측선택
      OR      M1504
      ANB
      AND=    K0 D3000
      MOV     K1 D3000
      MRD
      LD      D1021.4  ; 비금속 2층 좌측
      OR      D1021.A  ; 금속 2층 좌측
      ANB
      LD      M8013  ; 2층 좌측선택
      OR      M1504
      ANB
      AND=    K0 D3000
      MOV     K2 D3000
      MRD
      LD      D1021.1  ; 비금속 1층 우측
      OR      D1021.7  ; 금속 1층 우측
      ANB
      LD      M8010  ; 1층 우측 선택
      OR      M1504
      ANB
      AND=    K0 D3000
      MOV     K1 D3000
      MPP
      LD      D1021.2  ; 비금속 1층 좌측
      OR      D1021.8  ; 굼속1층 좌측
      ANB
      LD      M8011  ; 1층 좌측선택
      OR      M1504
      ANB
      AND=    K0 D3000
      MOV     K2 D3000
; 창고 전후진 완료
269   LD=     K1 D3000
      AND     X0D  ; 창고 후완
      MPS
      ANI     M1500
      SET     M550
      MPP
      LD      M1500
      OR      M1504
      ANB
      SET     M1501
281   LD=     K2 D3000
      AND     X0E  ; 창고 전완
      MPS
      ANI     M1500
      SET     M560
      MPP
      LD      M1500
      OR      M1504
      ANB
      SET     M1502
